(* IEC 61131-3 sources: PLC-Static-Analysis/modules/plc-rules/src/test/resources/PLCA-Q011, 2 files *)

(* ---- compliant.st ---- *)
FUNCTION_BLOCK FB_Ok
VAR_INPUT
    diPulses : DINT;
    rSpeed : REAL;
    nIn : INT;
END_VAR
VAR
    nPulses : INT;
    diWide : DINT;
    rOut : REAL;
    lrOut : LREAL;
    nUns : UINT;
    nSmall : SINT;
    bSel : BOOL;
END_VAR
VAR CONSTANT
    cLimit : DINT := 100;
END_VAR
nPulses := DINT_TO_INT(diPulses);
nPulses := nIn + 1;
nPulses := nIn * 2 + 7;
diWide := nIn;
rOut := rSpeed * 0.5;
rOut := nIn * 0.1;
lrOut := rSpeed;
nUns := nIn;
nSmall := 100;
rOut := nIn;
rOut := MAX(0.0, rSpeed);
nPulses := SEL(bSel, 102, 11);
nPulses := cLimit;
nUns := SIZEOF(rOut);
END_FUNCTION_BLOCK

(* ---- noncompliant.st ---- *)
FUNCTION_BLOCK FB_Count
VAR_INPUT
    diPulses : DINT;
    rSpeed : REAL;
    lrPos : LREAL;
    dwStatus : DWORD;
END_VAR
VAR
    nPulses : INT;
    nSpeed : INT;
    rPos : REAL;
    wStatus : WORD;
    nSmall : SINT;
    nUns : UINT;
END_VAR
nPulses := diPulses; // PLCA-Q011
nSpeed := rSpeed; // PLCA-Q011
rPos := lrPos; // PLCA-Q011
wStatus := dwStatus; // PLCA-Q011
nPulses := nPulses + diPulses; // PLCA-Q011
nSmall := 200; // PLCA-Q011
nUns := -1; // PLCA-Q011
F_Take(n := diPulses); // PLCA-Q011
F_Give(d => nPulses); // PLCA-Q011
END_FUNCTION_BLOCK

FUNCTION F_Take : BOOL
VAR_INPUT
    n : INT;
END_VAR
F_Take := n > 0;
END_FUNCTION

FUNCTION F_Give : BOOL
VAR_OUTPUT
    d : DINT;
END_VAR
d := 1;
END_FUNCTION
